// TIA Portal V21 export
TextList "TL_Kind"  ListRange=Decimal
  TextListEntry   Text="-"
  TextListEntry   From=1, To=1, Text="ISTOVAR Bay0->Bay1"
  TextListEntry   From=2, To=2, Text="UKRCAJ Bay1->Bay0"
